Staubli VAL3: stop.pgx

program stop()
// Lab2A Level 3 - shared manual simulation / physical cycle
begin
  // ============================================================
  // 1. REINICIAR EL CONTROL DE MOVIMIENTO
  // ============================================================
  resetMotion()

  // ============================================================
  // 2. PREPARAR LAS ORDENES DE PARADA
  // ============================================================
  // Parar el carro, ordenar que la barrera retenga
  // y dejar de soplar.
  trolleyOn = false
  barrierClosed = true
  blowOn = false

  // ============================================================
  // 3. SI ES FISICO, PARAR EL ADAPTADOR Y ESCRIBIR LAS SALIDAS
  // ============================================================
  if physicalRun
    taskKill("physicalIO")

    // Parar carro y soplado.
    io:bOut2 = false
    io:bOut1 = false

    // Retencion con la nueva polaridad: bOut5=0.
    // Debe coincidir con !barrierClosed del adaptador.
    io:bOut5 = false

    // No escribimos bOut0: conservamos la aspiracion.
    // Tampoco cambiamos aqui los actuadores de clasificacion.
  endIf


  // ============================================================
  // 4. INDICAR QUE SE HA EJECUTADO LA PARADA
  // ============================================================
  cycleStep = -1
  putln("Stopped - empty matrix before a new start")

end
